SUBAPPLICATION AUS_GT_0 (* Prüft ob USINT-Adapter Wert > 0 ist (AX-Adapter Ausgang) *)
  (* Standard: 61499-2 *)
  (* Version 1.0, 2026-10-15, franz, Meisterschulen am Ostbahnhof *)
  PACKAGE MyLib::sys;
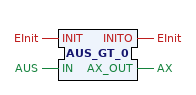
  EVENT_INPUT
    INIT : EInit; (* Initialization Request *)
  END_EVENT
  EVENT_OUTPUT
    INITO : EInit; (* Initialization Confirm *)
  END_EVENT
  SOCKETS
    IN : adapter::types::unidirectional::AUS;
  END_SOCKETS
  PLUGS
    AX_OUT : adapter::types::unidirectional::AX;
  END_PLUGS
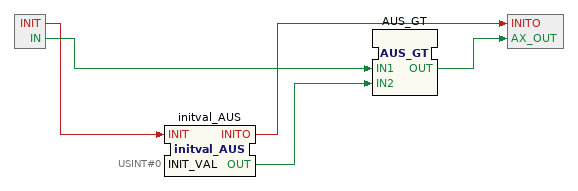
  FBS
    AUS_GT : adapter::iec61131::comparison::AUS_GT;
    initval_AUS : adapter::types::unidirectional::AUS::initval::initval_AUS(INIT_VAL := USINT#0);
  END_FBS
  EVENT_CONNECTIONS
    INIT TO initval_AUS.INIT;
    initval_AUS.INITO TO INITO;
  END_CONNECTIONS
  ADAPTER_CONNECTIONS
    IN TO AUS_GT.IN1;
    AUS_GT.OUT TO AX_OUT;
    initval_AUS.OUT TO AUS_GT.IN2;
  END_CONNECTIONS
END_SUBAPPLICATION
